(* IEC 61131-3 sources: model-first-plc-agent-ai/results/T2-B-27, 1 file *)

(* ---- b_code.st ---- *)
FUNCTION_BLOCK FillingControl
VAR_INPUT
    start : BOOL;
    stop : BOOL;
    LSH : BOOL;
    LSHH : BOOL;
    TimerDuration : TIME;
END_VAR
VAR_OUTPUT
    fill_valve : BOOL;
    discharge_valve : BOOL;
END_VAR
VAR
    current_step : INT := 0;
    filling_timer : TON;
    timer_done : BOOL := FALSE;
END_VAR

(* Stop and high-high level prevent entry into the filling step. *)
IF stop THEN
    current_step := 0;
ELSIF (current_step = 0) AND start AND NOT LSHH THEN
    current_step := 1;
END_IF;

filling_timer(
    IN := (current_step = 1) AND NOT stop AND NOT LSHH,
    PT := TimerDuration
);
timer_done := filling_timer.Q;

CASE current_step OF
    0:
        fill_valve := FALSE;

    1:
        IF stop OR LSHH OR timer_done THEN
            current_step := 0;
            fill_valve := FALSE;
        ELSE
            fill_valve := TRUE;
        END_IF;

ELSE
    current_step := 0;
    fill_valve := FALSE;
END_CASE;

discharge_valve := FALSE;

(* Reset immediately on leaving the filling step. *)
IF current_step = 0 THEN
    filling_timer(IN := FALSE, PT := TimerDuration);
END_IF;

END_FUNCTION_BLOCK

PROGRAM Main
VAR
    StartCommand AT %IX100.0 : BOOL;
    StopCommand AT %IX100.1 : BOOL;
    LSH AT %IX100.2 : BOOL;
    LSHH AT %IX100.3 : BOOL;
    FillValve AT %QX100.0 : BOOL;
    DischargeValve AT %QX100.1 : BOOL;
END_VAR
VAR
    TimerDuration : TIME := T#10s;
    start : BOOL := FALSE;
    stop : BOOL := FALSE;
    start_edge : R_TRIG;
    controller : FillingControl;
END_VAR

start_edge(CLK := StartCommand);
start := start_edge.Q;
stop := StopCommand;

controller(
    start := start,
    stop := stop,
    LSH := LSH,
    LSHH := LSHH,
    TimerDuration := TimerDuration
);

FillValve := controller.fill_valve;
DischargeValve := controller.discharge_valve;

END_PROGRAM
